(* IEC 61131-3 sources: plc_NativeGateway/src (part 3) *)

(* ---- NG_ReadAck.st ---- *)
FUNCTION_BLOCK NG_ReadAck
VAR_INPUT
    GatewayId : NG_Id;
END_VAR
VAR_IN_OUT
    Doc : NG_Document;
END_VAR
VAR_OUTPUT
    Valid : BOOL;
    MessageId : NG_Id;
    Stored : BOOL;
    Retryable : BOOL;
    Codes : NG_Text;
END_VAR
VAR
    RootFields : NG_AckFields;
    ErrorFields : NG_AckFields;
    t : INT;
    n : INT;
    e : INT;
    count : INT;
    code : NG_Text;
    wire : NG_Text;
END_VAR
Valid := FALSE; MessageId := ''; Stored := FALSE; Retryable := TRUE; Codes := '';
RootFields(Parent:=1,ErrorObject:=FALSE,Doc:=Doc); IF NOT RootFields.Valid THEN RETURN; END_IF;
t := RootFields.Fields[1]; IF (Doc.Tokens[t].Kind<>4) OR (Doc.Tokens[t].Number<>1) THEN RETURN; END_IF;
t := RootFields.Fields[2]; IF (Doc.Tokens[t].Kind<>3) OR (Doc.Tokens[t].Text<>GatewayId) THEN RETURN; END_IF;
t := RootFields.Fields[3];
(* Guard range before conversion. TO_LINT rounds and changes max-safe odd integers. *)
IF Doc.Tokens[t].Kind<>4 THEN RETURN; END_IF;
IF NOT ((Doc.Tokens[t].Number>=0) AND (Doc.Tokens[t].Number<=LREAL#9007199254740991.0)) THEN RETURN; END_IF;
IF Doc.Tokens[t].Number<>TO_LREAL(TRUNC_LINT(Doc.Tokens[t].Number)) THEN RETURN; END_IF;
t := RootFields.Fields[4];
IF (Doc.Tokens[t].Kind<>3) OR (LEN(Doc.Tokens[t].Text)>64) THEN RETURN; END_IF;
MessageId := Doc.Tokens[t].Text; IF NOT NG_ValidId(MessageId) THEN RETURN; END_IF;
t := RootFields.Fields[5]; IF Doc.Tokens[t].Kind<>3 THEN RETURN; END_IF;
IF Doc.Tokens[t].Text='STORED' THEN Stored:=TRUE;
ELSIF Doc.Tokens[t].Text<>'REJECTED' THEN RETURN; END_IF;
n := RootFields.Fields[6]; IF Doc.Tokens[n].Kind<>2 THEN RETURN; END_IF;
e:=n+1; count:=0;
WHILE e<Doc.Tokens[n].NextToken DO
    count:=count+1; IF Stored OR (count>32) THEN RETURN; END_IF;
    ErrorFields(Parent:=e,ErrorObject:=TRUE,Doc:=Doc); IF NOT ErrorFields.Valid THEN RETURN; END_IF;
    t:=ErrorFields.Fields[1]; IF (Doc.Tokens[t].Kind<>3) OR (Doc.Tokens[t].TextLength>256) THEN RETURN; END_IF;
    code:=Doc.Tokens[t].Text; wire:=NG_WireCode(code,FALSE); IF wire<>code THEN RETURN; END_IF;
    IF (code<>'UNKNOWN_CONFIG_VERSION') AND (code<>'RESOURCE_LIMIT') AND (code<>'STORAGE_ERROR') THEN Retryable:=FALSE; END_IF;
    IF LEN(Codes)<200 THEN IF Codes<>'' THEN Codes:=CONCAT(Codes,','); END_IF; Codes:=CONCAT(Codes,code); END_IF;
    t:=ErrorFields.Fields[2]; IF (Doc.Tokens[t].Kind<>3) OR (Doc.Tokens[t].TextLength>512) THEN RETURN; END_IF;
    IF (Doc.Tokens[t].Text<>'') AND (LEFT(Doc.Tokens[t].Text,1)<>'/') THEN RETURN; END_IF;
    t:=ErrorFields.Fields[3]; IF (Doc.Tokens[t].Kind<>3) OR (Doc.Tokens[t].TextLength<1) OR (Doc.Tokens[t].TextLength>256) THEN RETURN; END_IF;
    t:=ErrorFields.Fields[4];
    IF t>0 THEN IF (Doc.Tokens[t].Kind<>3) OR (LEN(Doc.Tokens[t].Text)>64) THEN RETURN; END_IF; wire:=Doc.Tokens[t].Text; IF NOT NG_ValidId(wire) THEN RETURN; END_IF; END_IF;
    t:=ErrorFields.Fields[5];
    IF t>0 THEN IF (Doc.Tokens[t].Kind<>3) OR (LEN(Doc.Tokens[t].Text)>64) THEN RETURN; END_IF; wire:=Doc.Tokens[t].Text; IF NOT NG_ValidId(wire) THEN RETURN; END_IF; END_IF;
    e:=Doc.Tokens[e].NextToken;
END_WHILE;
IF NOT Stored AND (count=0) THEN RETURN; END_IF;
Valid:=TRUE;
END_FUNCTION_BLOCK

(* ---- NG_ReadConfig.st ---- *)
FUNCTION_BLOCK NG_ReadConfig
VAR_INPUT
    Node : INT;
END_VAR
VAR_IN_OUT
    Doc : NG_Document;
    Config : NG_Config;
END_VAR
VAR_OUTPUT
    ErrorText : NG_Text;
END_VAR
VAR
    ReadDevice : NG_ReadDevice;
    Change : NG_EditDevice;
    Device : NG_Device;
    Points : ARRAY[1..32] OF NG_Point;
    t : INT;
    a : INT;
    d : INT;
    r : INT;
    err : NG_Text;
END_VAR
ErrorText := 'SCHEMA_INVALID';
IF NOT NG_Allowed(Node,'|enabled|report|devices|',Doc) THEN RETURN; END_IF;
t := NG_Member(Node,'enabled',Doc);
IF Doc.Tokens[t].Kind <> 5 THEN RETURN; END_IF;
Config.enabled := Doc.Tokens[t].Text = 'true';
r := NG_Member(Node,'report',Doc);
IF NOT NG_Allowed(r,'|batchIntervalMs|maxBatchPoints|',Doc) THEN RETURN; END_IF;
t := NG_Member(r,'batchIntervalMs',Doc);
IF (Doc.Tokens[t].Kind <> 4) OR (Doc.Tokens[t].Number < 1) OR (Doc.Tokens[t].Number > 86400000) OR (Doc.Tokens[t].Number <> TO_LREAL(TO_LINT(Doc.Tokens[t].Number))) THEN RETURN; END_IF;
Config.batchIntervalMs := TO_UDINT(Doc.Tokens[t].Number);
t := NG_Member(r,'maxBatchPoints',Doc);
IF (Doc.Tokens[t].Kind <> 4) OR (Doc.Tokens[t].Number < 1) OR (Doc.Tokens[t].Number > 500) OR (Doc.Tokens[t].Number <> TO_LREAL(TO_LINT(Doc.Tokens[t].Number))) THEN RETURN; END_IF;
Config.maxBatchPoints := TO_UINT(Doc.Tokens[t].Number);
a := NG_Member(Node,'devices',Doc);
IF Doc.Tokens[a].Kind <> 2 THEN RETURN; END_IF;
d := a + 1; Config.DeviceCount := 0; Config.PointCount := 0;
WHILE d < Doc.Tokens[a].NextToken DO
    IF Config.DeviceCount >= 50 THEN ErrorText := 'POINT_LIMIT_EXCEEDED'; RETURN; END_IF;
    ReadDevice(Node := d, Doc := Doc, Device := Device, Points := Points);
    err := ReadDevice.ErrorText;
    IF err <> '' THEN ErrorText := err; RETURN; END_IF;
    Change(DeviceIndex := Config.DeviceCount+1, Remove := FALSE, Replacement := Device, Config := Config, Points := Points);
    IF Change.ErrorText <> '' THEN ErrorText := Change.ErrorText; RETURN; END_IF;
    d := Doc.Tokens[d].NextToken;
END_WHILE;
ErrorText := NG_CheckConfig(Config);
END_FUNCTION_BLOCK

(* ---- NG_ReadDevice.st ---- *)
FUNCTION_BLOCK NG_ReadDevice
VAR_INPUT
    Node : INT;
END_VAR
VAR_IN_OUT
    Doc : NG_Document;
    Device : NG_Device;
    Points : ARRAY[1..32] OF NG_Point;
END_VAR
VAR_OUTPUT
    ErrorText : NG_Text;
END_VAR
VAR
    ReadPoint : NG_ReadPoint;
    t : INT;
    conn : INT;
    pointsNode : INT;
    p : INT;
    err : NG_Text;
END_VAR
ErrorText := '';
IF NOT NG_Allowed(Node,'|deviceId|name|enabled|protocol|connection|points|',Doc) THEN ErrorText := 'SCHEMA_INVALID'; RETURN; END_IF;
t := NG_Member(Node, 'deviceId', Doc);
IF (Doc.Tokens[t].Kind <> 3) OR (LEN(Doc.Tokens[t].Text) < 1) OR (LEN(Doc.Tokens[t].Text) > 64) THEN ErrorText := 'SCHEMA_INVALID'; RETURN; END_IF;
Device.deviceId := Doc.Tokens[t].Text;
t := NG_Member(Node, 'name', Doc);
IF (Doc.Tokens[t].Kind <> 3) OR (LEN(Doc.Tokens[t].Text) < 1) OR (LEN(Doc.Tokens[t].Text) > 128) THEN ErrorText := 'SCHEMA_INVALID'; RETURN; END_IF;
Device.name := Doc.Tokens[t].Text;
t := NG_Member(Node, 'enabled', Doc);
IF (Doc.Tokens[t].Kind <> 5) THEN ErrorText := 'SCHEMA_INVALID'; RETURN; END_IF;
Device.enabled := (Doc.Tokens[t].Text = 'true');
t := NG_Member(Node,'protocol',Doc);
IF (Doc.Tokens[t].Kind <> 3) OR (Doc.Tokens[t].Text <> 'modbus_tcp') THEN ErrorText := 'UNSUPPORTED_PROTOCOL'; RETURN; END_IF;
conn := NG_Member(Node,'connection',Doc);
IF NOT NG_Allowed(conn,'|host|port|unitId|connectTimeoutMs|requestTimeoutMs|retryCount|maxReadRegisters|maxRegisterGap|',Doc) THEN ErrorText := 'SCHEMA_INVALID'; RETURN; END_IF;
t := NG_Member(conn, 'host', Doc);
IF (Doc.Tokens[t].Kind <> 3) OR (LEN(Doc.Tokens[t].Text) < 1) OR (LEN(Doc.Tokens[t].Text) > 253) THEN ErrorText := 'SCHEMA_INVALID'; RETURN; END_IF;
Device.host := Doc.Tokens[t].Text;
t := NG_Member(conn, 'port', Doc);
IF (Doc.Tokens[t].Kind <> 4) OR (Doc.Tokens[t].Number < LREAL#1.0) OR (Doc.Tokens[t].Number > LREAL#65535.0) OR (Doc.Tokens[t].Number <> TO_LREAL(TO_LINT(Doc.Tokens[t].Number))) THEN ErrorText := 'SCHEMA_INVALID'; RETURN; END_IF;
Device.port := TO_UINT(Doc.Tokens[t].Number);
t := NG_Member(conn, 'unitId', Doc);
IF (Doc.Tokens[t].Kind <> 4) OR (Doc.Tokens[t].Number < LREAL#0.0) OR (Doc.Tokens[t].Number > LREAL#255.0) OR (Doc.Tokens[t].Number <> TO_LREAL(TO_LINT(Doc.Tokens[t].Number))) THEN ErrorText := 'SCHEMA_INVALID'; RETURN; END_IF;
Device.unitId := TO_USINT(Doc.Tokens[t].Number);
t := NG_Member(conn, 'connectTimeoutMs', Doc);
IF (Doc.Tokens[t].Kind <> 4) OR (Doc.Tokens[t].Number < LREAL#1.0) OR (Doc.Tokens[t].Number > LREAL#300000.0) OR (Doc.Tokens[t].Number <> TO_LREAL(TO_LINT(Doc.Tokens[t].Number))) THEN ErrorText := 'SCHEMA_INVALID'; RETURN; END_IF;
Device.connectTimeoutMs := TO_UDINT(Doc.Tokens[t].Number);
t := NG_Member(conn, 'requestTimeoutMs', Doc);
IF (Doc.Tokens[t].Kind <> 4) OR (Doc.Tokens[t].Number < LREAL#1.0) OR (Doc.Tokens[t].Number > LREAL#300000.0) OR (Doc.Tokens[t].Number <> TO_LREAL(TO_LINT(Doc.Tokens[t].Number))) THEN ErrorText := 'SCHEMA_INVALID'; RETURN; END_IF;
Device.requestTimeoutMs := TO_UDINT(Doc.Tokens[t].Number);
t := NG_Member(conn, 'retryCount', Doc);
IF (Doc.Tokens[t].Kind <> 4) OR (Doc.Tokens[t].Number < LREAL#0.0) OR (Doc.Tokens[t].Number > LREAL#10.0) OR (Doc.Tokens[t].Number <> TO_LREAL(TO_LINT(Doc.Tokens[t].Number))) THEN ErrorText := 'SCHEMA_INVALID'; RETURN; END_IF;
Device.retryCount := TO_USINT(Doc.Tokens[t].Number);
t := NG_Member(conn, 'maxReadRegisters', Doc);
IF t > 0 THEN
    IF (Doc.Tokens[t].Kind <> 4) OR (Doc.Tokens[t].Number < LREAL#1.0) OR (Doc.Tokens[t].Number > LREAL#125.0) OR (Doc.Tokens[t].Number <> TO_LREAL(TO_LINT(Doc.Tokens[t].Number))) THEN ErrorText := 'SCHEMA_INVALID'; RETURN; END_IF;
    Device.maxReadRegisters := TO_UINT(Doc.Tokens[t].Number);
ELSE
    Device.maxReadRegisters := UINT#0;
END_IF;
t := NG_Member(conn, 'maxRegisterGap', Doc);
IF t > 0 THEN
    IF (Doc.Tokens[t].Kind <> 4) OR (Doc.Tokens[t].Number < LREAL#0.0) OR (Doc.Tokens[t].Number > LREAL#124.0) OR (Doc.Tokens[t].Number <> TO_LREAL(TO_LINT(Doc.Tokens[t].Number))) THEN ErrorText := 'SCHEMA_INVALID'; RETURN; END_IF;
    Device.hasMaxRegisterGap := TRUE;
    Device.maxRegisterGap := TO_UINT(Doc.Tokens[t].Number);
ELSE
    Device.hasMaxRegisterGap := FALSE;
    Device.maxRegisterGap := UINT#0;
END_IF;
pointsNode := NG_Member(Node,'points',Doc);
IF Doc.Tokens[pointsNode].Kind <> 2 THEN ErrorText := 'SCHEMA_INVALID'; RETURN; END_IF;
Device.PointCount := 0; p := pointsNode + 1;
WHILE p < Doc.Tokens[pointsNode].NextToken DO
    IF Device.PointCount >= 32 THEN ErrorText := 'POINT_LIMIT_EXCEEDED'; RETURN; END_IF;
    Device.PointCount := Device.PointCount + 1;
    ReadPoint(Node := p, Doc := Doc, Point := Points[Device.PointCount]);
    err := ReadPoint.ErrorText;
    IF err <> '' THEN ErrorText := err; RETURN; END_IF;
    p := Doc.Tokens[p].NextToken;
END_WHILE;

END_FUNCTION_BLOCK

(* ---- NG_ReadPoint.st ---- *)
FUNCTION_BLOCK NG_ReadPoint
VAR_INPUT
    Node : INT;
END_VAR
VAR_IN_OUT
    Doc : NG_Document;
    Point : NG_Point;
END_VAR
VAR_OUTPUT
    ErrorText : NG_Text;
END_VAR
VAR
    t : INT;
    mb : INT;
END_VAR
ErrorText := '';
IF NOT NG_Allowed(Node,'|pointId|name|enabled|dataType|pollIntervalMs|scale|offset|unit|reportMode|reportIntervalMs|deadband|staleAfterMs|modbus|',Doc) THEN ErrorText := 'SCHEMA_INVALID'; RETURN; END_IF;
t := NG_Member(Node, 'pointId', Doc);
IF (Doc.Tokens[t].Kind <> 3) OR (LEN(Doc.Tokens[t].Text) < 1) OR (LEN(Doc.Tokens[t].Text) > 64) THEN ErrorText := 'SCHEMA_INVALID'; RETURN; END_IF;
Point.pointId := Doc.Tokens[t].Text;
t := NG_Member(Node, 'name', Doc);
IF (Doc.Tokens[t].Kind <> 3) OR (LEN(Doc.Tokens[t].Text) < 1) OR (LEN(Doc.Tokens[t].Text) > 128) THEN ErrorText := 'SCHEMA_INVALID'; RETURN; END_IF;
Point.name := Doc.Tokens[t].Text;
t := NG_Member(Node, 'enabled', Doc);
IF (Doc.Tokens[t].Kind <> 5) THEN ErrorText := 'SCHEMA_INVALID'; RETURN; END_IF;
Point.enabled := (Doc.Tokens[t].Text = 'true');
t := NG_Member(Node, 'dataType', Doc);
IF (Doc.Tokens[t].Kind <> 3) OR (LEN(Doc.Tokens[t].Text) < 1) OR (LEN(Doc.Tokens[t].Text) > 16) THEN ErrorText := 'SCHEMA_INVALID'; RETURN; END_IF;
Point.dataType := Doc.Tokens[t].Text;
t := NG_Member(Node, 'pollIntervalMs', Doc);
IF (Doc.Tokens[t].Kind <> 4) OR (Doc.Tokens[t].Number < LREAL#1.0) OR (Doc.Tokens[t].Number > LREAL#86400000.0) OR (Doc.Tokens[t].Number <> TO_LREAL(TO_LINT(Doc.Tokens[t].Number))) THEN ErrorText := 'SCHEMA_INVALID'; RETURN; END_IF;
Point.pollIntervalMs := TO_UDINT(Doc.Tokens[t].Number);
t := NG_Member(Node, 'scale', Doc);
IF (Doc.Tokens[t].Kind <> 4) OR (Doc.Tokens[t].Number < LREAL#-1.0E+100) OR (Doc.Tokens[t].Number > LREAL#1.0E+100) THEN ErrorText := 'SCHEMA_INVALID'; RETURN; END_IF;
Point.scale := Doc.Tokens[t].Number;
t := NG_Member(Node, 'offset', Doc);
IF (Doc.Tokens[t].Kind <> 4) OR (Doc.Tokens[t].Number < LREAL#-1.0E+100) OR (Doc.Tokens[t].Number > LREAL#1.0E+100) THEN ErrorText := 'SCHEMA_INVALID'; RETURN; END_IF;
Point.offset := Doc.Tokens[t].Number;
t := NG_Member(Node, 'unit', Doc);
IF t > 0 THEN
IF (Doc.Tokens[t].Kind <> 3) OR (LEN(Doc.Tokens[t].Text) < 0) OR (LEN(Doc.Tokens[t].Text) > 32) THEN ErrorText := 'SCHEMA_INVALID'; RETURN; END_IF;
Point.unit := Doc.Tokens[t].Text;
ELSE Point.unit := ''; END_IF;
t := NG_Member(Node, 'reportMode', Doc);
IF (Doc.Tokens[t].Kind <> 3) OR (LEN(Doc.Tokens[t].Text) < 1) OR (LEN(Doc.Tokens[t].Text) > 24) THEN ErrorText := 'SCHEMA_INVALID'; RETURN; END_IF;
Point.reportMode := Doc.Tokens[t].Text;
t := NG_Member(Node, 'reportIntervalMs', Doc);
IF (Doc.Tokens[t].Kind <> 4) OR (Doc.Tokens[t].Number < LREAL#1.0) OR (Doc.Tokens[t].Number > LREAL#86400000.0) OR (Doc.Tokens[t].Number <> TO_LREAL(TO_LINT(Doc.Tokens[t].Number))) THEN ErrorText := 'SCHEMA_INVALID'; RETURN; END_IF;
Point.reportIntervalMs := TO_UDINT(Doc.Tokens[t].Number);
t := NG_Member(Node, 'deadband', Doc);
IF (Doc.Tokens[t].Kind <> 4) OR (Doc.Tokens[t].Number < LREAL#0.0) OR (Doc.Tokens[t].Number > LREAL#1.0E+100) THEN ErrorText := 'SCHEMA_INVALID'; RETURN; END_IF;
Point.deadband := Doc.Tokens[t].Number;
t := NG_Member(Node, 'staleAfterMs', Doc);
IF (Doc.Tokens[t].Kind <> 4) OR (Doc.Tokens[t].Number < LREAL#1.0) OR (Doc.Tokens[t].Number > LREAL#86400000.0) OR (Doc.Tokens[t].Number <> TO_LREAL(TO_LINT(Doc.Tokens[t].Number))) THEN ErrorText := 'SCHEMA_INVALID'; RETURN; END_IF;
Point.staleAfterMs := TO_UDINT(Doc.Tokens[t].Number);
mb := NG_Member(Node,'modbus',Doc);
IF NOT NG_Allowed(mb,'|area|address|byteOrder|',Doc) THEN ErrorText := 'SCHEMA_INVALID'; RETURN; END_IF;
t := NG_Member(mb, 'area', Doc);
IF (Doc.Tokens[t].Kind <> 3) OR (LEN(Doc.Tokens[t].Text) < 1) OR (LEN(Doc.Tokens[t].Text) > 24) THEN ErrorText := 'SCHEMA_INVALID'; RETURN; END_IF;
Point.area := Doc.Tokens[t].Text;
t := NG_Member(mb, 'address', Doc);
IF (Doc.Tokens[t].Kind <> 4) OR (Doc.Tokens[t].Number < LREAL#0.0) OR (Doc.Tokens[t].Number > LREAL#65535.0) OR (Doc.Tokens[t].Number <> TO_LREAL(TO_LINT(Doc.Tokens[t].Number))) THEN ErrorText := 'SCHEMA_INVALID'; RETURN; END_IF;
Point.address := TO_UINT(Doc.Tokens[t].Number);
t := NG_Member(mb, 'byteOrder', Doc);
IF t > 0 THEN
IF (Doc.Tokens[t].Kind <> 3) OR (LEN(Doc.Tokens[t].Text) < 0) OR (LEN(Doc.Tokens[t].Text) > 4) THEN ErrorText := 'SCHEMA_INVALID'; RETURN; END_IF;
Point.byteOrder := Doc.Tokens[t].Text;
ELSE Point.byteOrder := ''; END_IF;
END_FUNCTION_BLOCK

(* ---- NG_ReportPolicy.st ---- *)
FUNCTION_BLOCK NG_ReportPolicy
VAR_INPUT
    DeferCapacity : BOOL;
END_VAR
VAR_IN_OUT
    Buffer : NG_Buffer;
END_VAR
VAR
    Event : NG_CaptureEvent;
    Gap : NG_GapLog;
    AuditDecision : NG_AuditDecision;
    s : UINT;
    p : UINT;
    r : UINT;
    c : UINT;
    n : INT;
    slots : ULINT;
    selected : BOOL;
    present : BOOL;
    reject : BOOL;
    reason : USINT;
END_VAR

(* Atomic RAM admission is this mode's local commit boundary. The copied
   baseline has no dependency on delivery order or subsequent slot reuse. *)
FOR n:=1 TO 64 DO
    IF Buffer.WorkDeadlineUs>0 THEN IF GET_MICROSECONDS(TRUE)+ULINT#70>=Buffer.WorkDeadlineUs THEN EXIT; END_IF; END_IF;
    IF Buffer.IngressCount=0 THEN EXIT; END_IF;
    (* A local whole-batch reclaim may need the next bounded scan. Keep this
       raw event undecided until that reclaim; never wait on SDK/ACK here. *)
    IF DeferCapacity AND (Buffer.FreeHead=0) AND (Buffer.HighSlot>=28800) THEN EXIT; END_IF;
    Event:=Buffer.Ingress[Buffer.Head]; s:=Event.ConfigSlot; p:=Event.PointIndex;
    Buffer.Head:=Buffer.Head MOD 512+1; Buffer.IngressCount:=Buffer.IngressCount-1;
    reject:=FALSE; reason:=0;
    IF (s<>Buffer.ActiveSlot) OR (Event.ConfigGeneration<>Buffer.Configs[s].Generation) OR
       (Event.SamplingGeneration<>Buffer.SamplingGeneration) OR NOT Buffer.Cursors[p].Enabled THEN
        Buffer.UndecidedLostEventsTotal:=NG_SafeAdd(Buffer.UndecidedLostEventsTotal,ULINT#1);
        Buffer.AccountingComplete:=FALSE;
        reason:=2; reject:=TRUE;
    ELSE
        present:=((Event.Flags AND WORD#1)<>WORD#0) AND
                 (((Event.Flags AND WORD#2)<>WORD#0) OR ((Event.Flags AND WORD#8)<>WORD#0));
        IF Buffer.PlatformTime THEN
            present:=present AND Buffer.TimeValid AND (Event.ClockRevision=Buffer.ClockRevision)
                AND ((Event.Flags AND WORD#2)<>WORD#0);
        END_IF;
        IF (Buffer.ReportCursors[p].SamplingGeneration<>Event.SamplingGeneration) OR
           (Buffer.ReportCursors[p].ConfigGeneration<>Event.ConfigGeneration) OR
           (Buffer.ReportCursors[p].ClockRevision<>Event.ClockRevision) OR
           (Buffer.ReportCursors[p].TimePresent<>present) THEN
            slots:=Buffer.Cursors[p].ActivatedMonoMs;
            IF (Buffer.ReportCursors[p].ConfigGeneration=Event.ConfigGeneration) AND
               ((Buffer.ReportCursors[p].TimePresent<>present) OR (Buffer.ReportCursors[p].ClockRevision<>Event.ClockRevision)) THEN
                slots:=Buffer.Cursors[p].NextDueMonoMs;
                IF Event.Kind=1 THEN slots:=Event.NominalDueMonoMs; END_IF;
            END_IF;
            Buffer.ReportCursors[p].SamplingGeneration:=Event.SamplingGeneration;
            Buffer.ReportCursors[p].ConfigGeneration:=Event.ConfigGeneration;
            Buffer.ReportCursors[p].ClockRevision:=Event.ClockRevision;
            Buffer.ReportCursors[p].TimePresent:=present;
            Buffer.ReportCursors[p].HasBaseline:=FALSE;
            Buffer.ReportCursors[p].NextDue:=slots;
        END_IF;
        selected:=NOT Buffer.ReportCursors[p].HasBaseline OR (Buffer.ReportCursors[p].Quality<>Event.Quality);
        IF Buffer.ReportCursors[p].HasBaseline AND (Event.Quality=2) AND (Buffer.ReportCursors[p].Quality=2) AND
           (Buffer.Configs[s].Config.Points[p].reportMode<>'cyclic') THEN
            IF Buffer.Configs[s].Config.Points[p].dataType='bool' THEN
                selected:=selected OR ((Event.Value=LREAL#0.0)<>(Buffer.ReportCursors[p].Value=LREAL#0.0));
            ELSE selected:=selected OR (ABS(Event.Value-Buffer.ReportCursors[p].Value)>Buffer.Configs[s].Config.Points[p].deadband); END_IF;
        END_IF;
        IF (Event.Kind=1) AND (Buffer.Configs[s].Config.Points[p].reportMode<>'change') AND
           (Event.NominalDueMonoMs>=Buffer.ReportCursors[p].NextDue) THEN
            slots:=(Event.NominalDueMonoMs-Buffer.ReportCursors[p].NextDue)/TO_ULINT(Buffer.Configs[s].Config.Points[p].reportIntervalMs)+1;
            Buffer.MissedReportSlotsTotal:=NG_SafeAdd(Buffer.MissedReportSlotsTotal,slots-1);
            Buffer.ReportCursors[p].NextDue:=Buffer.ReportCursors[p].NextDue+slots*TO_ULINT(Buffer.Configs[s].Config.Points[p].reportIntervalMs);
            selected:=TRUE;
        END_IF;
        IF NOT selected THEN
            Buffer.PolicyFilteredEventsTotal:=NG_SafeAdd(Buffer.PolicyFilteredEventsTotal,ULINT#1); reject:=TRUE;
        ELSE
            Buffer.EligibleEventsTotal:=NG_SafeAdd(Buffer.EligibleEventsTotal,ULINT#1);
            IF NOT present THEN
                Buffer.TimeInvalidEventsTotal:=NG_SafeAdd(Buffer.TimeInvalidEventsTotal,ULINT#1); reason:=4; reject:=TRUE;
            ELSIF (Buffer.FreeHead=0) AND (Buffer.HighSlot>=28800) THEN
                Buffer.EnqueueRejectedAttemptsTotal:=NG_SafeAdd(Buffer.EnqueueRejectedAttemptsTotal,ULINT#1); reason:=5; reject:=TRUE;
            END_IF;
            IF reject THEN Buffer.KnownUnsentEventsTotal:=NG_SafeAdd(Buffer.KnownUnsentEventsTotal,ULINT#1); END_IF;
        END_IF;
    END_IF;
    IF reject THEN
        c:=1;
        IF reason=2 THEN c:=4; ELSIF reason<>0 THEN c:=3; END_IF;
        AuditDecision(SampleSeq:=Event.SampleSeq,Decision:=TO_USINT(c),Reason:=reason,Buffer:=Buffer);
        IF reason<>0 THEN Gap(Reason:=reason,Event:=Event,Buffer:=Buffer); END_IF;
        Buffer.Configs[s].References:=Buffer.Configs[s].References-1;
    ELSE
        IF Buffer.FreeHead<>0 THEN r:=Buffer.FreeHead; Buffer.FreeHead:=Buffer.FreeSlots[r];
        ELSE Buffer.HighSlot:=Buffer.HighSlot+1; r:=Buffer.HighSlot; END_IF;
        IF Buffer.RecordGenerations[r]=UDINT#4294967295 THEN Buffer.CaptureStopped:=TRUE;
            Buffer.KnownUnsentEventsTotal:=NG_SafeAdd(Buffer.KnownUnsentEventsTotal,ULINT#1);
            Gap(Reason:=USINT#5,Event:=Event,Buffer:=Buffer); Buffer.Configs[s].References:=Buffer.Configs[s].References-1;
            AuditDecision(SampleSeq:=Event.SampleSeq,Decision:=USINT#3,Reason:=USINT#5,Buffer:=Buffer);
        ELSE
            Buffer.RecordGenerations[r]:=Buffer.RecordGenerations[r]+1;
            Buffer.Records[r]:=Event; Buffer.RecordStates[r]:=1; Buffer.FreeSlots[r]:=0;
            Buffer.LastAdmittedSeq:=MAX(Buffer.LastAdmittedSeq,Event.SampleSeq);
            AuditDecision(SampleSeq:=Event.SampleSeq,Decision:=USINT#2,Reason:=USINT#0,Buffer:=Buffer);
            Buffer.OwnedCount:=Buffer.OwnedCount+1;
            c:=2; IF Event.SampleSeq<=Buffer.Watermark THEN c:=1; END_IF;
            IF Buffer.QueueHead[c]=0 THEN Buffer.QueueHead[c]:=r; ELSE Buffer.FreeSlots[Buffer.QueueTail[c]]:=r; END_IF;
            Buffer.QueueTail[c]:=r;
            IF Event.SampleSeq>Buffer.ReportCursors[p].LastSeq THEN
                Buffer.ReportCursors[p].LastSeq:=Event.SampleSeq; Buffer.ReportCursors[p].Value:=Event.Value;
                Buffer.ReportCursors[p].Quality:=Event.Quality; Buffer.ReportCursors[p].HasBaseline:=TRUE;
            END_IF;
        END_IF;
    END_IF;
END_FOR;
END_FUNCTION_BLOCK

(* ---- NG_Resources.st ---- *)
FUNCTION_BLOCK NG_Resources
VAR_INPUT
    NowMs : ULINT;
END_VAR
VAR_OUTPUT
    Changed : BOOL;
    MemoryValid : BOOL;
    CpuValid : BOOL;
    ProcessValid : BOOL;
    TotalKiB : ULINT;
    AvailableKiB : ULINT;
    RssKiB : ULINT;
    CpuPermille : UDINT;
    ProcessName : STRING[64];
    ErrorText : NG_Text;
END_VAR
VAR
    OpenFile : FILE_OPEN;
    ReadFile : FILE_READ;
    CloseFile : FILE_CLOSE;
    Convert : BUF_TO_STRING;
    Name : STRING;
    Bytes : NG_ProcBytes;
    Text : NG_ProcText;
    Stage : INT;
    FileIndex : INT := 1;
    Handle : UINT;
    Count : UDINT;
    NextRead : ULINT;
    p : INT;
    c : INT;
    n : INT;
    start : INT;
    token : ULINT;
    total : ULINT;
    idle : ULINT;
    PrevTotal : ULINT;
    PrevIdle : ULINT;
    HasDigit : BOOL;
    ProcFailed : BOOL;
END_VAR
Changed := FALSE;
CASE FileIndex OF
1: Name := '/proc/meminfo';
2: Name := '/proc/stat';
3: Name := '/proc/self/status';
END_CASE;
OpenFile(Execute := Stage=10, Name := Name);
ReadFile(Execute := Stage=20, Handle := Handle, MaxLength := UDINT#8191, Buffer := Bytes);
CloseFile(Execute := Stage=30, Handle := Handle);
Convert(REQ := Stage=40, BUF_FORMAT := FALSE, BUF_OFFS := 0, BUF_CNT := TO_INT(Count), BUFFER := Bytes, DST := Text);
CASE Stage OF
0:
    IF NowMs >= NextRead THEN FileIndex := 1; ErrorText := ''; ProcFailed := FALSE; Stage := 10; END_IF;
10:
    IF OpenFile.Error THEN ProcFailed := TRUE; Stage := 80;
    ELSIF OpenFile.Done THEN Handle := OpenFile.Handle; Stage := 20; END_IF;
20:
    IF ReadFile.Error OR ReadFile.Done THEN Count := ReadFile.LengthRead; ProcFailed := Count=0; Stage := 30; END_IF;
30:
    IF CloseFile.Done OR CloseFile.Error THEN IF CloseFile.Error OR ProcFailed THEN Stage := 80; ELSE Stage := 40; END_IF; END_IF;
40:
    IF Convert.ERROR THEN ProcFailed := TRUE; Stage := 80;
    ELSIF Convert.DONE THEN
        CASE FileIndex OF
        1:
            TotalKiB := NG_ProcNumber(Text,'MemTotal:'); AvailableKiB := NG_ProcNumber(Text,'MemAvailable:');
            IF AvailableKiB=0 THEN AvailableKiB := NG_ProcNumber(Text,'MemFree:')+NG_ProcNumber(Text,'Buffers:')+NG_ProcNumber(Text,'Cached:'); END_IF;
            MemoryValid := TotalKiB > 0;
        2:
            total := 0; idle := 0; n := 0; token := 0; HasDigit := FALSE;
            p := FIND(Text,'cpu ');
            IF p > 0 THEN
                p := p+4;
                WHILE p <= LEN(Text) DO
                    c := GET_CHAR(Text,p);
                    IF (c>=48) AND (c<=57) THEN token := token*10+TO_ULINT(c-48); HasDigit := TRUE;
                    ELSE
                        IF HasDigit THEN
                            n := n+1; IF n <= 8 THEN total := total+token; END_IF;
                            IF (n=4) OR (n=5) THEN idle := idle+token; END_IF;
                            token := 0; HasDigit := FALSE;
                        END_IF;
                        IF (c=10) OR (n>=8) THEN EXIT; END_IF;
                    END_IF;
                    p := p+1;
                END_WHILE;
                IF (PrevTotal > 0) AND (total > PrevTotal) AND (idle >= PrevIdle) THEN
                    CpuPermille := TO_UDINT((total-PrevTotal-(idle-PrevIdle))*1000/(total-PrevTotal)); CpuValid := TRUE;
                END_IF;
                PrevTotal := total; PrevIdle := idle;
            END_IF;
        3:
            RssKiB := NG_ProcNumber(Text,'VmRSS:'); ProcessValid := RssKiB > 0;
            start := FIND(Text,'Name:');
            IF start > 0 THEN
                start := start+5;
                WHILE start <= LEN(Text) DO c := GET_CHAR(Text,start); IF (c<>32) AND (c<>9) THEN EXIT; END_IF; start := start+1; END_WHILE;
                p := start;
                WHILE p <= LEN(Text) DO IF GET_CHAR(Text,p)=10 THEN EXIT; END_IF; p := p+1; END_WHILE;
                IF p > start THEN ProcessName := MID(Text,MIN(63,p-start),start); END_IF;
            END_IF;
        END_CASE;
        Stage := 80;
    END_IF;
80:
    IF ProcFailed THEN
        ErrorText := CONCAT('PROC_READ_FAILED:',TO_STRING(FileIndex,'{0:d}'));
        CASE FileIndex OF 1: MemoryValid := FALSE; 2: CpuValid := FALSE; 3: ProcessValid := FALSE; END_CASE;
    END_IF;
    ProcFailed := FALSE;
    IF FileIndex < 3 THEN FileIndex := FileIndex+1; Stage := 10;
    ELSE Changed := TRUE; NextRead := NowMs+10000; Stage := 0; END_IF;
END_CASE;
END_FUNCTION_BLOCK

(* ---- NG_SameConfig.st ---- *)
FUNCTION_BLOCK NG_SameConfig
VAR_OUTPUT
    Equal : BOOL;
END_VAR
VAR_IN_OUT
    A : NG_Config;
    B : NG_Config;
END_VAR
VAR
    i : INT;
END_VAR
Equal := FALSE;
IF (A.Version<>B.Version) OR (A.MessageId<>B.MessageId) OR (A.enabled<>B.enabled) OR
   (A.batchIntervalMs<>B.batchIntervalMs) OR (A.maxBatchPoints<>B.maxBatchPoints) OR
   (A.DeviceCount<>B.DeviceCount) OR (A.PointCount<>B.PointCount) THEN RETURN; END_IF;
FOR i:=1 TO A.DeviceCount DO
    IF (A.Devices[i].deviceId<>B.Devices[i].deviceId) OR (A.Devices[i].name<>B.Devices[i].name) OR
       (A.Devices[i].enabled<>B.Devices[i].enabled) OR (A.Devices[i].host<>B.Devices[i].host) OR
       (A.Devices[i].port<>B.Devices[i].port) OR (A.Devices[i].unitId<>B.Devices[i].unitId) OR
       (A.Devices[i].connectTimeoutMs<>B.Devices[i].connectTimeoutMs) OR
       (A.Devices[i].requestTimeoutMs<>B.Devices[i].requestTimeoutMs) OR
       (A.Devices[i].retryCount<>B.Devices[i].retryCount) OR
       (A.Devices[i].maxReadRegisters<>B.Devices[i].maxReadRegisters) OR
       (A.Devices[i].hasMaxRegisterGap<>B.Devices[i].hasMaxRegisterGap) OR
       (A.Devices[i].maxRegisterGap<>B.Devices[i].maxRegisterGap) OR
       (A.Devices[i].PointStart<>B.Devices[i].PointStart) OR (A.Devices[i].PointCount<>B.Devices[i].PointCount) THEN RETURN; END_IF;
END_FOR;
FOR i:=1 TO A.PointCount DO
    IF (A.Points[i].pointId<>B.Points[i].pointId) OR (A.Points[i].name<>B.Points[i].name) OR
       (A.Points[i].enabled<>B.Points[i].enabled) OR (A.Points[i].dataType<>B.Points[i].dataType) OR
       (A.Points[i].pollIntervalMs<>B.Points[i].pollIntervalMs) OR (A.Points[i].scale<>B.Points[i].scale) OR
       (A.Points[i].offset<>B.Points[i].offset) OR (A.Points[i].unit<>B.Points[i].unit) OR
       (A.Points[i].reportMode<>B.Points[i].reportMode) OR (A.Points[i].reportIntervalMs<>B.Points[i].reportIntervalMs) OR
       (A.Points[i].deadband<>B.Points[i].deadband) OR (A.Points[i].staleAfterMs<>B.Points[i].staleAfterMs) OR
       (A.Points[i].area<>B.Points[i].area) OR (A.Points[i].address<>B.Points[i].address) OR
       (A.Points[i].byteOrder<>B.Points[i].byteOrder) THEN RETURN; END_IF;
END_FOR;
Equal := TRUE;
END_FUNCTION_BLOCK

(* ---- NG_SHA256.st ---- *)
FUNCTION_BLOCK NG_SHA256
VAR_INPUT
    Execute : BOOL;
    Length : UDINT;
END_VAR
VAR_IN_OUT
    Buffer : NG_Bytes;
END_VAR
VAR_OUTPUT
    Busy : BOOL;
    Done : BOOL;
    Digest : STRING[64];
END_VAR
VAR
    Prev : BOOL;
    Block : UDINT;
    Blocks : UDINT;
    Offset : UDINT;
    i : INT;
    j : INT;
    n : INT;
    v : DWORD;
    a : DWORD;
    b : DWORD;
    c : DWORD;
    d : DWORD;
    e : DWORD;
    f : DWORD;
    g : DWORD;
    h : DWORD;
    s0 : DWORD;
    s1 : DWORD;
    t1 : DWORD;
    t2 : DWORD;
    Hs : ARRAY[0..7] OF DWORD;
    W : ARRAY[0..63] OF DWORD;
    K : ARRAY[0..63] OF DWORD := [16#428A2F98,16#71374491,16#B5C0FBCF,16#E9B5DBA5,16#3956C25B,16#59F111F1,16#923F82A4,16#AB1C5ED5,16#D807AA98,16#12835B01,16#243185BE,16#550C7DC3,16#72BE5D74,16#80DEB1FE,16#9BDC06A7,16#C19BF174,16#E49B69C1,16#EFBE4786,16#0FC19DC6,16#240CA1CC,16#2DE92C6F,16#4A7484AA,16#5CB0A9DC,16#76F988DA,16#983E5152,16#A831C66D,16#B00327C8,16#BF597FC7,16#C6E00BF3,16#D5A79147,16#06CA6351,16#14292967,16#27B70A85,16#2E1B2138,16#4D2C6DFC,16#53380D13,16#650A7354,16#766A0ABB,16#81C2C92E,16#92722C85,16#A2BFE8A1,16#A81A664B,16#C24B8B70,16#C76C51A3,16#D192E819,16#D6990624,16#F40E3585,16#106AA070,16#19A4C116,16#1E376C08,16#2748774C,16#34B0BCB5,16#391C0CB3,16#4ED8AA4A,16#5B9CCA4F,16#682E6FF3,16#748F82EE,16#78A5636F,16#84C87814,16#8CC70208,16#90BEFFFA,16#A4506CEB,16#BEF9A3F7,16#C67178F2];
END_VAR
IF Execute AND NOT Prev AND NOT Busy THEN
    Hs[0] := 16#6A09E667; Hs[1] := 16#BB67AE85; Hs[2] := 16#3C6EF372; Hs[3] := 16#A54FF53A;
    Hs[4] := 16#510E527F; Hs[5] := 16#9B05688C; Hs[6] := 16#1F83D9AB; Hs[7] := 16#5BE0CD19;
    Block := 0; Blocks := (Length + 72) / 64; Busy := TRUE; Done := FALSE; Digest := '';
END_IF;
Prev := Execute;
IF NOT Busy THEN RETURN; END_IF;
FOR n := 1 TO 8 DO
    FOR i := 0 TO 15 DO
        W[i] := 0;
        FOR j := 0 TO 3 DO
            Offset := Block*64 + TO_UDINT(i*4+j);
            IF Offset < Length THEN v := TO_DWORD(Buffer[Offset]);
            ELSIF Offset = Length THEN v := DWORD#16#80;
            ELSIF Offset >= Blocks*64-8 THEN v := TO_DWORD(SHR(TO_LWORD(TO_ULINT(Length)*ULINT#8),TO_UINT((Blocks*64-1-Offset)*8)) AND LWORD#255);
            ELSE v := 0; END_IF;
            W[i] := SHL(W[i],8) OR v;
        END_FOR;
    END_FOR;
    FOR i := 16 TO 63 DO
        s0 := ROR(W[i-15],7) XOR ROR(W[i-15],18) XOR SHR(W[i-15],3);
        s1 := ROR(W[i-2],17) XOR ROR(W[i-2],19) XOR SHR(W[i-2],10);
        W[i] := NG_Add4(W[i-16],s0,W[i-7],s1);
    END_FOR;
    a := Hs[0]; b := Hs[1]; c := Hs[2]; d := Hs[3]; e := Hs[4]; f := Hs[5]; g := Hs[6]; h := Hs[7];
    FOR i := 0 TO 63 DO
        s1 := ROR(e,6) XOR ROR(e,11) XOR ROR(e,25);
        t1 := NG_Add4(h,s1,(e AND f) XOR ((NOT e) AND g),K[i]);
        t1 := NG_Add4(t1,W[i],DWORD#0,DWORD#0);
        s0 := ROR(a,2) XOR ROR(a,13) XOR ROR(a,22);
        t2 := NG_Add4(s0,(a AND b) XOR (a AND c) XOR (b AND c),DWORD#0,DWORD#0);
        h := g; g := f; f := e; e := NG_Add4(d,t1,DWORD#0,DWORD#0);
        d := c; c := b; b := a; a := NG_Add4(t1,t2,DWORD#0,DWORD#0);
    END_FOR;
    Hs[0] := NG_Add4(Hs[0],a,DWORD#0,DWORD#0); Hs[1] := NG_Add4(Hs[1],b,DWORD#0,DWORD#0);
    Hs[2] := NG_Add4(Hs[2],c,DWORD#0,DWORD#0); Hs[3] := NG_Add4(Hs[3],d,DWORD#0,DWORD#0);
    Hs[4] := NG_Add4(Hs[4],e,DWORD#0,DWORD#0); Hs[5] := NG_Add4(Hs[5],f,DWORD#0,DWORD#0);
    Hs[6] := NG_Add4(Hs[6],g,DWORD#0,DWORD#0); Hs[7] := NG_Add4(Hs[7],h,DWORD#0,DWORD#0);
    Block := Block + 1;
    IF Block >= Blocks THEN
        FOR i := 0 TO 7 DO Digest := CONCAT(Digest,TO_STRING(Hs[i],'{0:x8}')); END_FOR;
        Busy := FALSE; Done := TRUE; EXIT;
    END_IF;
END_FOR;
END_FUNCTION_BLOCK

(* ---- NG_SourceResult.st ---- *)
FUNCTION_BLOCK NG_SourceResult
VAR_INPUT
    Index : UINT;
    Value : LREAL;
    Quality : STRING[24];
    NowMs : ULINT;
    UnixMs : ULINT;
    NominalDueMs : ULINT;
    ConfigSlot : UINT;
    ConfigGeneration : UDINT;
    SamplingGeneration : ULINT;
END_VAR
VAR_OUTPUT
    Accepted : BOOL;
END_VAR
VAR_IN_OUT
    Samples : ARRAY[1..320] OF NG_Sample;
    Buffer : NG_Buffer;
END_VAR
VAR
    Core : NG_SourceResultCore;
END_VAR
(* Bind each bounded source/sample/deadline once for the final physical result. *)
Accepted:=FALSE;
IF (Index<1) OR (Index>320) THEN RETURN; END_IF;
Core(Index:=Index,Value:=Value,Quality:=Quality,NowMs:=NowMs,UnixMs:=UnixMs,NominalDueMs:=NominalDueMs,ConfigSlot:=ConfigSlot,ConfigGeneration:=ConfigGeneration,SamplingGeneration:=SamplingGeneration,Cursor:=Buffer.Cursors[Index],Sample:=Samples[Index],StaleDue:=Buffer.SourceStaleDue[Index],Buffer:=Buffer);
Accepted:=Core.Accepted;
END_FUNCTION_BLOCK

(* ---- NG_SourceResultCore.st ---- *)
FUNCTION_BLOCK NG_SourceResultCore
VAR_INPUT
    Index : UINT;
    Value : LREAL;
    Quality : STRING[24];
    NowMs : ULINT;
    UnixMs : ULINT;
    NominalDueMs : ULINT;
    ConfigSlot : UINT;
    ConfigGeneration : UDINT;
    SamplingGeneration : ULINT;
END_VAR
VAR_OUTPUT
    Accepted : BOOL;
END_VAR
VAR_IN_OUT
    Cursor : NG_SourceCursor;
    Sample : NG_Sample;
    StaleDue : ULINT;
    Buffer : NG_Buffer;
END_VAR
VAR
    Capture : NG_Capture;
    code : USINT;
    text : STRING[24];
END_VAR
Accepted:=FALSE;
IF (Index<1) OR (Index>320) OR (ConfigSlot=0) OR (ConfigSlot>4) THEN RETURN; END_IF;
IF (ConfigSlot<>Buffer.ActiveSlot) OR (Buffer.Configs[ConfigSlot].Generation<>ConfigGeneration) OR
   (Buffer.SamplingGeneration<>SamplingGeneration) OR NOT Cursor.Enabled THEN
    Buffer.CancelledReadsTotal:=NG_SafeAdd(Buffer.CancelledReadsTotal,ULINT#1);
    Buffer.CancellationReason:=2; RETURN;
END_IF;
IF NowMs<NominalDueMs THEN Buffer.CaptureStopped:=TRUE; RETURN; END_IF;
text:=Quality;
IF (text='GOOD') AND NOT (ABS(Value)<=LREAL#1.7976931348623157E308) THEN text:='BAD_DECODE'; END_IF;
code:=NG_QualityCode(text);
Capture(PointIndex:=Index, Kind:=USINT#1, Quality:=code, Value:=Value, NowMs:=NowMs, NominalDueMs:=NominalDueMs, SystemUtcMs:=UnixMs, Buffer:=Buffer);
    Accepted:=Capture.Accepted;
Cursor.LastPhysicalMonoMs:=NowMs; Cursor.HasPhysical:=TRUE;
Cursor.Quality:=code;
(* A final result extends this source's liveness. Keeping an earlier global
   deadline is safe; the due sweep recomputes the minimum before emitting stale. *)
StaleDue:=0;
IF code<>3 THEN
    StaleDue:=NowMs+TO_ULINT(Buffer.Configs[ConfigSlot].Config.Points[Index].staleAfterMs);
    IF StaleDue<Buffer.StaleCheckAt THEN Buffer.StaleCheckAt:=StaleDue; END_IF;
END_IF;
Sample.Quality:=text; Sample.Timestamp:=UnixMs; Sample.Fresh:=TRUE;
IF text='GOOD' THEN Sample.Value:=Value; Sample.LastGoodMs:=NowMs; END_IF;
Sample.NextPollMs:=Cursor.NextDueMonoMs;
END_FUNCTION_BLOCK

(* ---- NG_SourceState.st ---- *)
FUNCTION_BLOCK NG_SourceState
VAR_INPUT
    Index : UINT;
    Enabled : BOOL;
    NowMs : ULINT;
    UnixMs : ULINT;
    StaleAfterMs : UDINT;
    CheckStale : BOOL;
END_VAR
VAR_OUTPUT
    Accepted : BOOL;
END_VAR
VAR_IN_OUT
    Samples : ARRAY[1..320] OF NG_Sample;
    Buffer : NG_Buffer;
END_VAR
VAR
    Core : NG_SourceStateCore;
END_VAR
(* Bind each bounded source/sample reference once. Repeated field updates in
   Core avoid dozens of generated array-bound helper calls per activation. *)
Accepted:=FALSE;
IF (Index<1) OR (Index>320) THEN RETURN; END_IF;
Core(Index:=Index,Enabled:=Enabled,NowMs:=NowMs,UnixMs:=UnixMs,
    StaleAfterMs:=StaleAfterMs,CheckStale:=CheckStale,
    Cursor:=Buffer.Cursors[Index],Sample:=Samples[Index],Buffer:=Buffer);
Accepted:=Core.Accepted;
END_FUNCTION_BLOCK

(* ---- NG_SourceStateCore.st ---- *)
FUNCTION_BLOCK NG_SourceStateCore
VAR_INPUT
    Index : UINT;
    Enabled : BOOL;
    NowMs : ULINT;
    UnixMs : ULINT;
    StaleAfterMs : UDINT;
    CheckStale : BOOL;
END_VAR
VAR_OUTPUT
    Accepted : BOOL;
END_VAR
VAR_IN_OUT
    Cursor : NG_SourceCursor;
    Sample : NG_Sample;
    Buffer : NG_Buffer;
END_VAR
VAR
    Capture : NG_CaptureCore;
    start : ULINT;
END_VAR

Accepted:=FALSE;
IF (Index<1) OR (Index>320) THEN RETURN; END_IF;
IF NOT Enabled THEN Cursor.Enabled:=FALSE; Buffer.SourceStaleDue[Index]:=0; RETURN; END_IF;
IF (Cursor.Generation<>Buffer.SamplingGeneration) OR NOT Cursor.Enabled THEN
    Cursor.Generation:=Buffer.SamplingGeneration; Cursor.Enabled:=TRUE;
    Cursor.ActivatedMonoMs:=NowMs; Cursor.LastPhysicalMonoMs:=0;
    Cursor.HasPhysical:=FALSE; Cursor.HasPhysicalUtc:=FALSE;
    Cursor.NextDueMonoMs:=NowMs; Cursor.Quality:=1;
    Buffer.SourceStaleDue[Index]:=NowMs+TO_ULINT(StaleAfterMs);
    IF Buffer.SourceStaleDue[Index]<Buffer.StaleCheckAt THEN Buffer.StaleCheckAt:=Buffer.SourceStaleDue[Index]; END_IF;
    Sample.Quality:='UNKNOWN'; Sample.Timestamp:=UnixMs; Sample.Fresh:=TRUE;
    Sample.NextPollMs:=NowMs;
    Capture(PointIndex:=Index, Kind:=USINT#2, Quality:=USINT#1, Value:=LREAL#0.0, NowMs:=NowMs, NominalDueMs:=ULINT#0, SystemUtcMs:=UnixMs, Cursor:=Cursor, Buffer:=Buffer);
    Accepted:=Capture.Accepted;
END_IF;
IF NOT CheckStale THEN RETURN; END_IF;
start:=Cursor.ActivatedMonoMs;
IF Cursor.HasPhysical THEN start:=Cursor.LastPhysicalMonoMs; END_IF;
IF (NowMs>=start) AND (NowMs-start>=TO_ULINT(StaleAfterMs)) AND (Cursor.Quality<>3) THEN
    Cursor.Quality:=3; Sample.Quality:='STALE';
    Buffer.SourceStaleDue[Index]:=0;
    Sample.Timestamp:=UnixMs; Sample.Fresh:=TRUE;
    Capture(PointIndex:=Index, Kind:=USINT#2, Quality:=USINT#3, Value:=LREAL#0.0, NowMs:=NowMs, NominalDueMs:=ULINT#0, SystemUtcMs:=UnixMs, Cursor:=Cursor, Buffer:=Buffer);
    Accepted:=Capture.Accepted;
END_IF;
END_FUNCTION_BLOCK

(* ---- NG_StorageHash.st ---- *)
FUNCTION_BLOCK NG_StorageHash
VAR_INPUT
    Execute : BOOL;
    Length : UDINT;
END_VAR
VAR_IN_OUT
    Buffer : NG_StorageBytes;
END_VAR
VAR_OUTPUT
    Busy : BOOL;
    Done : BOOL;
    Digest : STRING[64];
END_VAR
VAR
    Prev : BOOL;
    Block : UDINT;
    Blocks : UDINT;
    Offset : UDINT;
    i : INT;
    j : INT;
    n : INT;
    v : DWORD;
    a : DWORD;
    b : DWORD;
    c : DWORD;
    d : DWORD;
    e : DWORD;
    f : DWORD;
    g : DWORD;
    h : DWORD;
    s0 : DWORD;
    s1 : DWORD;
    t1 : DWORD;
    t2 : DWORD;
    Hs : ARRAY[0..7] OF DWORD;
    W : ARRAY[0..63] OF DWORD;
    K : ARRAY[0..63] OF DWORD := [16#428A2F98,16#71374491,16#B5C0FBCF,16#E9B5DBA5,16#3956C25B,16#59F111F1,16#923F82A4,16#AB1C5ED5,16#D807AA98,16#12835B01,16#243185BE,16#550C7DC3,16#72BE5D74,16#80DEB1FE,16#9BDC06A7,16#C19BF174,16#E49B69C1,16#EFBE4786,16#0FC19DC6,16#240CA1CC,16#2DE92C6F,16#4A7484AA,16#5CB0A9DC,16#76F988DA,16#983E5152,16#A831C66D,16#B00327C8,16#BF597FC7,16#C6E00BF3,16#D5A79147,16#06CA6351,16#14292967,16#27B70A85,16#2E1B2138,16#4D2C6DFC,16#53380D13,16#650A7354,16#766A0ABB,16#81C2C92E,16#92722C85,16#A2BFE8A1,16#A81A664B,16#C24B8B70,16#C76C51A3,16#D192E819,16#D6990624,16#F40E3585,16#106AA070,16#19A4C116,16#1E376C08,16#2748774C,16#34B0BCB5,16#391C0CB3,16#4ED8AA4A,16#5B9CCA4F,16#682E6FF3,16#748F82EE,16#78A5636F,16#84C87814,16#8CC70208,16#90BEFFFA,16#A4506CEB,16#BEF9A3F7,16#C67178F2];
END_VAR
IF Execute AND NOT Prev AND NOT Busy THEN
    Hs[0] := 16#6A09E667; Hs[1] := 16#BB67AE85; Hs[2] := 16#3C6EF372; Hs[3] := 16#A54FF53A;
    Hs[4] := 16#510E527F; Hs[5] := 16#9B05688C; Hs[6] := 16#1F83D9AB; Hs[7] := 16#5BE0CD19;
    Block := 0; Blocks := (Length + 72) / 64; Busy := TRUE; Done := FALSE; Digest := '';
END_IF;
Prev := Execute;
IF NOT Busy THEN RETURN; END_IF;
FOR n := 1 TO 16 DO
    FOR i := 0 TO 15 DO
        W[i] := 0;
        FOR j := 0 TO 3 DO
            Offset := Block*64 + TO_UDINT(i*4+j);
            IF Offset < Length THEN v := TO_DWORD(Buffer[Offset]);
            ELSIF Offset = Length THEN v := DWORD#16#80;
            ELSIF Offset >= Blocks*64-8 THEN v := TO_DWORD(SHR(TO_LWORD(TO_ULINT(Length)*ULINT#8),TO_UINT((Blocks*64-1-Offset)*8)) AND LWORD#255);
            ELSE v := 0; END_IF;
            W[i] := SHL(W[i],8) OR v;
        END_FOR;
    END_FOR;
    FOR i := 16 TO 63 DO
        s0 := ROR(W[i-15],7) XOR ROR(W[i-15],18) XOR SHR(W[i-15],3);
        s1 := ROR(W[i-2],17) XOR ROR(W[i-2],19) XOR SHR(W[i-2],10);
        W[i] := NG_Add4(W[i-16],s0,W[i-7],s1);
    END_FOR;
    a := Hs[0]; b := Hs[1]; c := Hs[2]; d := Hs[3]; e := Hs[4]; f := Hs[5]; g := Hs[6]; h := Hs[7];
    FOR i := 0 TO 63 DO
        s1 := ROR(e,6) XOR ROR(e,11) XOR ROR(e,25);
        t1 := NG_Add4(h,s1,(e AND f) XOR ((NOT e) AND g),K[i]);
        t1 := NG_Add4(t1,W[i],DWORD#0,DWORD#0);
        s0 := ROR(a,2) XOR ROR(a,13) XOR ROR(a,22);
        t2 := NG_Add4(s0,(a AND b) XOR (a AND c) XOR (b AND c),DWORD#0,DWORD#0);
        h := g; g := f; f := e; e := NG_Add4(d,t1,DWORD#0,DWORD#0);
        d := c; c := b; b := a; a := NG_Add4(t1,t2,DWORD#0,DWORD#0);
    END_FOR;
    Hs[0] := NG_Add4(Hs[0],a,DWORD#0,DWORD#0); Hs[1] := NG_Add4(Hs[1],b,DWORD#0,DWORD#0);
    Hs[2] := NG_Add4(Hs[2],c,DWORD#0,DWORD#0); Hs[3] := NG_Add4(Hs[3],d,DWORD#0,DWORD#0);
    Hs[4] := NG_Add4(Hs[4],e,DWORD#0,DWORD#0); Hs[5] := NG_Add4(Hs[5],f,DWORD#0,DWORD#0);
    Hs[6] := NG_Add4(Hs[6],g,DWORD#0,DWORD#0); Hs[7] := NG_Add4(Hs[7],h,DWORD#0,DWORD#0);
    Block := Block + 1;
    IF Block >= Blocks THEN
        FOR i := 0 TO 7 DO Digest := CONCAT(Digest,TO_STRING(Hs[i],'{0:x8}')); END_FOR;
        Busy := FALSE; Done := TRUE; EXIT;
    END_IF;
END_FOR;
END_FUNCTION_BLOCK

(* ---- NG_Store.st ---- *)
FUNCTION_BLOCK NG_Store
VAR_INPUT
    Save : BOOL;
END_VAR
VAR_IN_OUT
    Candidate : NG_Durable;
END_VAR
VAR_OUTPUT
    Ready : BOOL;
    NeedsMigration : BOOL;
    Busy : BOOL;
    Done : BOOL;
    Error : BOOL;
    ErrorText : NG_Text;
    Active : NG_Durable;
END_VAR
VAR
    LegacyRecord : NG1_File;
    V2Record : NG2_File;
    V3Record : NG3_File;
    V4Record : NG4_File;
    V4 : BOOL;
    V3 : BOOL;
    V2 : BOOL;
    Legacy : BOOL;
    StateLength : UDINT;
    d : INT;
    p : INT;
    idx : INT;
    Stage : INT;
    Slot : INT := 1;
    ActiveSlot : INT;
    Prev : BOOL;
    Name : STRING;
    OpenFile : FILE_OPEN;
    ReadFile : FILE_READ;
    WriteFile : FILE_WRITE;
    CloseFile : FILE_CLOSE;
    Handle : UINT;
    Record : NG_File;
    Verify : NG_File;
    Bytes : NG_StorageBytes;
    CopyBytes : BUF_TO_BYTE;
    Hash : NG_StorageHash;
    Valid : BOOL;
    Saving : BOOL;
    OperationFailed : BOOL;
END_VAR
Done := FALSE;
IF Legacy THEN
    IF Slot = 1 THEN Name := '/opt/plcnext/NativeGateway-A.bin'; ELSE Name := '/opt/plcnext/NativeGateway-B.bin'; END_IF;
    StateLength := SIZEOF(LegacyRecord.State);
ELSIF V2 THEN
    IF Slot = 1 THEN Name := '/opt/plcnext/NativeGateway-v2-A.bin'; ELSE Name := '/opt/plcnext/NativeGateway-v2-B.bin'; END_IF;
    StateLength := SIZEOF(V2Record.State);
ELSIF V3 THEN
    IF Slot = 1 THEN Name := '/opt/plcnext/NativeGateway-v3-A.bin'; ELSE Name := '/opt/plcnext/NativeGateway-v3-B.bin'; END_IF;
    StateLength := SIZEOF(V3Record.State);
ELSIF V4 THEN
    IF Slot = 1 THEN Name := '/opt/plcnext/NativeGateway-v4-A.bin'; ELSE Name := '/opt/plcnext/NativeGateway-v4-B.bin'; END_IF;
    StateLength := SIZEOF(V4Record.State);
ELSE
    IF Slot = 1 THEN Name := '/opt/plcnext/NativeGateway-v5-A.bin'; ELSE Name := '/opt/plcnext/NativeGateway-v5-B.bin'; END_IF;
    StateLength := SIZEOF(Record.State);
END_IF;
OpenFile(Execute := (Stage = 10) OR (Stage = 60) OR (Stage = 90), Name := Name);
IF Legacy THEN
    ReadFile(Execute := Stage = 20, Handle := Handle, MaxLength := SIZEOF(LegacyRecord), Buffer := LegacyRecord);
ELSIF V2 THEN
    ReadFile(Execute := Stage = 20, Handle := Handle, MaxLength := SIZEOF(V2Record), Buffer := V2Record);
ELSIF V3 THEN
    ReadFile(Execute := Stage = 20, Handle := Handle, MaxLength := SIZEOF(V3Record), Buffer := V3Record);
ELSIF V4 THEN
    ReadFile(Execute := Stage = 20, Handle := Handle, MaxLength := SIZEOF(V4Record), Buffer := V4Record);
ELSE
    ReadFile(Execute := (Stage = 20) OR (Stage = 100), Handle := Handle, MaxLength := SIZEOF(Record), Buffer := Record);
END_IF;
WriteFile(Execute := Stage = 70, Handle := Handle, Length := SIZEOF(Record), Buffer := Record);
CloseFile(Execute := (Stage = 30) OR (Stage = 80) OR (Stage = 110) OR (Stage = 900), Handle := Handle);
IF Legacy THEN
    CopyBytes(REQ := Stage = 35, BUF_FORMAT := FALSE, BUF_OFFS := 0, BUF_CNT := StateLength, BUFFER := LegacyRecord.State, DST := Bytes);
ELSIF V2 THEN
    CopyBytes(REQ := Stage = 35, BUF_FORMAT := FALSE, BUF_OFFS := 0, BUF_CNT := StateLength, BUFFER := V2Record.State, DST := Bytes);
ELSIF V3 THEN
    CopyBytes(REQ := Stage = 35, BUF_FORMAT := FALSE, BUF_OFFS := 0, BUF_CNT := StateLength, BUFFER := V3Record.State, DST := Bytes);
ELSIF V4 THEN
    CopyBytes(REQ := Stage = 35, BUF_FORMAT := FALSE, BUF_OFFS := 0, BUF_CNT := StateLength, BUFFER := V4Record.State, DST := Bytes);
ELSE
    CopyBytes(REQ := (Stage = 35) OR (Stage = 50) OR (Stage = 115), BUF_FORMAT := FALSE, BUF_OFFS := 0, BUF_CNT := StateLength, BUFFER := Record.State, DST := Bytes);
END_IF;
Hash(Execute := (Stage = 40) OR (Stage = 55) OR (Stage = 120), Length := StateLength, Buffer := Bytes);
CASE Stage OF
0: Ready := FALSE; Busy := TRUE; Slot := 1; Stage := 10;
10:
    IF OpenFile.Error THEN Stage := 45;
    ELSIF OpenFile.Done THEN Handle := OpenFile.Handle; Stage := 20;
    END_IF;
20:
    IF ReadFile.Error OR ReadFile.Done THEN
        IF Legacy THEN Valid := ReadFile.Done AND (ReadFile.LengthRead = SIZEOF(LegacyRecord)) AND (LegacyRecord.Magic = DWORD#16#4E475731) AND (LegacyRecord.FormatVersion = 1);
        ELSIF V2 THEN Valid := ReadFile.Done AND (ReadFile.LengthRead = SIZEOF(V2Record)) AND (V2Record.Magic = DWORD#16#4E475732) AND (V2Record.FormatVersion = 2);
        ELSIF V3 THEN Valid := ReadFile.Done AND (ReadFile.LengthRead = SIZEOF(V3Record)) AND (V3Record.Magic = DWORD#16#4E475733) AND (V3Record.FormatVersion = 3);
        ELSIF V4 THEN Valid := ReadFile.Done AND (ReadFile.LengthRead = SIZEOF(V4Record)) AND (V4Record.Magic = DWORD#16#4E475734) AND (V4Record.FormatVersion = 4);
        ELSE Valid := ReadFile.Done AND (ReadFile.LengthRead = SIZEOF(Record)) AND (Record.Magic = DWORD#16#4E475735) AND (Record.FormatVersion = 5); END_IF;
        Stage := 30;
    END_IF;
30:
    IF CloseFile.Done OR CloseFile.Error THEN
        IF Valid AND NOT CloseFile.Error THEN Stage := 35; ELSE Stage := 45; END_IF;
    END_IF;
35: IF CopyBytes.DONE THEN Stage := 40; ELSIF CopyBytes.ERROR THEN Stage := 45; END_IF;
40:
    IF Hash.Done THEN
        IF Legacy THEN
            IF (Hash.Digest = LegacyRecord.Digest) AND (LegacyRecord.State.Generation > Active.Generation) THEN
                Active.Managed := FALSE; Active.BootCounter := 0;
                Active.Generation := LegacyRecord.State.Generation; Active.Bootstrap := LegacyRecord.State.Bootstrap;
                Active.ReplayIndex := LegacyRecord.State.ReplayIndex; Active.Requests := LegacyRecord.State.Requests;
                Active.Config.Version := LegacyRecord.State.Config.Version; Active.Config.MessageId := LegacyRecord.State.Config.MessageId;
                Active.Config.enabled := LegacyRecord.State.Config.enabled; Active.Config.batchIntervalMs := LegacyRecord.State.Config.batchIntervalMs;
                Active.Config.maxBatchPoints := LegacyRecord.State.Config.maxBatchPoints; Active.Config.DeviceCount := LegacyRecord.State.Config.DeviceCount;
                idx := 1;
                FOR d := 1 TO Active.Config.DeviceCount DO
                    Active.Config.Devices[d].deviceId := LegacyRecord.State.Config.Devices[d].deviceId;
                    Active.Config.Devices[d].name := LegacyRecord.State.Config.Devices[d].name;
                    Active.Config.Devices[d].enabled := LegacyRecord.State.Config.Devices[d].enabled;
                    Active.Config.Devices[d].host := LegacyRecord.State.Config.Devices[d].host;
                    Active.Config.Devices[d].port := LegacyRecord.State.Config.Devices[d].port;
                    Active.Config.Devices[d].unitId := LegacyRecord.State.Config.Devices[d].unitId;
                    Active.Config.Devices[d].connectTimeoutMs := LegacyRecord.State.Config.Devices[d].connectTimeoutMs;
                    Active.Config.Devices[d].requestTimeoutMs := LegacyRecord.State.Config.Devices[d].requestTimeoutMs;
                    Active.Config.Devices[d].retryCount := LegacyRecord.State.Config.Devices[d].retryCount;
                    Active.Config.Devices[d].maxReadRegisters := UINT#0;
                    Active.Config.Devices[d].hasMaxRegisterGap := FALSE;
                    Active.Config.Devices[d].maxRegisterGap := UINT#0;
                    Active.Config.Devices[d].PointCount := LegacyRecord.State.Config.Devices[d].PointCount;
                    Active.Config.Devices[d].PointStart := idx;
                    FOR p := 1 TO Active.Config.Devices[d].PointCount DO Active.Config.Points[idx] := LegacyRecord.State.Config.Devices[d].Points[p]; idx := idx+1; END_FOR;
                END_FOR;
                Active.Config.PointCount := idx-1; NeedsMigration := TRUE;
            END_IF;
        ELSIF V2 THEN
            IF (Hash.Digest = V2Record.Digest) AND (V2Record.State.Generation > Active.Generation) THEN
                Active.Generation := V2Record.State.Generation; Active.Bootstrap := V2Record.State.Bootstrap;
                Active.Config.Version := V2Record.State.Config.Version; Active.Config.MessageId := V2Record.State.Config.MessageId;
                Active.Config.enabled := V2Record.State.Config.enabled; Active.Config.batchIntervalMs := V2Record.State.Config.batchIntervalMs;
                Active.Config.maxBatchPoints := V2Record.State.Config.maxBatchPoints; Active.Config.DeviceCount := V2Record.State.Config.DeviceCount;
                Active.Config.PointCount := V2Record.State.Config.PointCount; Active.Config.Points := V2Record.State.Config.Points;
                FOR d := 1 TO Active.Config.DeviceCount DO
                    Active.Config.Devices[d].deviceId := V2Record.State.Config.Devices[d].deviceId; Active.Config.Devices[d].name := V2Record.State.Config.Devices[d].name;
                    Active.Config.Devices[d].enabled := V2Record.State.Config.Devices[d].enabled; Active.Config.Devices[d].host := V2Record.State.Config.Devices[d].host;
                    Active.Config.Devices[d].port := V2Record.State.Config.Devices[d].port; Active.Config.Devices[d].unitId := V2Record.State.Config.Devices[d].unitId;
                    Active.Config.Devices[d].connectTimeoutMs := V2Record.State.Config.Devices[d].connectTimeoutMs; Active.Config.Devices[d].requestTimeoutMs := V2Record.State.Config.Devices[d].requestTimeoutMs;
                    Active.Config.Devices[d].retryCount := V2Record.State.Config.Devices[d].retryCount;
                    Active.Config.Devices[d].maxReadRegisters := UINT#0; Active.Config.Devices[d].hasMaxRegisterGap := FALSE; Active.Config.Devices[d].maxRegisterGap := UINT#0;
                    Active.Config.Devices[d].PointCount := V2Record.State.Config.Devices[d].PointCount; Active.Config.Devices[d].PointStart := V2Record.State.Config.Devices[d].PointStart;
                END_FOR;
                Active.Requests := V2Record.State.Requests; Active.ReplayIndex := V2Record.State.ReplayIndex;
                Active.Managed := FALSE; Active.BootCounter := 0; NeedsMigration := TRUE;
            END_IF;
        ELSIF V3 THEN
            IF (Hash.Digest = V3Record.Digest) AND (V3Record.State.Generation > Active.Generation) THEN
                Active.Generation := V3Record.State.Generation; Active.Managed := V3Record.State.Managed;
                Active.BootCounter := V3Record.State.BootCounter; Active.Bootstrap := V3Record.State.Bootstrap;
                Active.Config.Version := V3Record.State.Config.Version; Active.Config.MessageId := V3Record.State.Config.MessageId;
                Active.Config.enabled := V3Record.State.Config.enabled; Active.Config.batchIntervalMs := V3Record.State.Config.batchIntervalMs;
                Active.Config.maxBatchPoints := V3Record.State.Config.maxBatchPoints; Active.Config.DeviceCount := V3Record.State.Config.DeviceCount;
                Active.Config.PointCount := V3Record.State.Config.PointCount; Active.Config.Points := V3Record.State.Config.Points;
                FOR d := 1 TO Active.Config.DeviceCount DO
                    Active.Config.Devices[d].deviceId := V3Record.State.Config.Devices[d].deviceId; Active.Config.Devices[d].name := V3Record.State.Config.Devices[d].name;
                    Active.Config.Devices[d].enabled := V3Record.State.Config.Devices[d].enabled; Active.Config.Devices[d].host := V3Record.State.Config.Devices[d].host;
                    Active.Config.Devices[d].port := V3Record.State.Config.Devices[d].port; Active.Config.Devices[d].unitId := V3Record.State.Config.Devices[d].unitId;
                    Active.Config.Devices[d].connectTimeoutMs := V3Record.State.Config.Devices[d].connectTimeoutMs; Active.Config.Devices[d].requestTimeoutMs := V3Record.State.Config.Devices[d].requestTimeoutMs;
                    Active.Config.Devices[d].retryCount := V3Record.State.Config.Devices[d].retryCount;
                    Active.Config.Devices[d].maxReadRegisters := UINT#0; Active.Config.Devices[d].hasMaxRegisterGap := FALSE; Active.Config.Devices[d].maxRegisterGap := UINT#0;
                    Active.Config.Devices[d].PointCount := V3Record.State.Config.Devices[d].PointCount; Active.Config.Devices[d].PointStart := V3Record.State.Config.Devices[d].PointStart;
                END_FOR;
                Active.Requests := V3Record.State.Requests; Active.ReplayIndex := V3Record.State.ReplayIndex;
                Active.HasHubBaseline := Active.Managed AND (Active.Config.Version > 0);
                IF Active.HasHubBaseline THEN Active.HubConfig := Active.Config; END_IF;
                Active.LocalChanges := FALSE; Active.LocalRevision := 0; NeedsMigration := TRUE;
            END_IF;
        ELSIF V4 THEN
            IF (Hash.Digest = V4Record.Digest) AND (V4Record.State.Generation > Active.Generation) THEN
                Active.Generation := V4Record.State.Generation; Active.Managed := V4Record.State.Managed;
                Active.BootCounter := V4Record.State.BootCounter; Active.Bootstrap := V4Record.State.Bootstrap;
                Active.HasHubBaseline := V4Record.State.HasHubBaseline; Active.LocalChanges := V4Record.State.LocalChanges; Active.LocalRevision := V4Record.State.LocalRevision;
                Active.Config.Version := V4Record.State.Config.Version; Active.Config.MessageId := V4Record.State.Config.MessageId;
                Active.Config.enabled := V4Record.State.Config.enabled; Active.Config.batchIntervalMs := V4Record.State.Config.batchIntervalMs;
                Active.Config.maxBatchPoints := V4Record.State.Config.maxBatchPoints; Active.Config.DeviceCount := V4Record.State.Config.DeviceCount;
                Active.Config.PointCount := V4Record.State.Config.PointCount; Active.Config.Points := V4Record.State.Config.Points;
                FOR d := 1 TO Active.Config.DeviceCount DO
                    Active.Config.Devices[d].deviceId := V4Record.State.Config.Devices[d].deviceId; Active.Config.Devices[d].name := V4Record.State.Config.Devices[d].name;
                    Active.Config.Devices[d].enabled := V4Record.State.Config.Devices[d].enabled; Active.Config.Devices[d].host := V4Record.State.Config.Devices[d].host;
                    Active.Config.Devices[d].port := V4Record.State.Config.Devices[d].port; Active.Config.Devices[d].unitId := V4Record.State.Config.Devices[d].unitId;
                    Active.Config.Devices[d].connectTimeoutMs := V4Record.State.Config.Devices[d].connectTimeoutMs; Active.Config.Devices[d].requestTimeoutMs := V4Record.State.Config.Devices[d].requestTimeoutMs;
                    Active.Config.Devices[d].retryCount := V4Record.State.Config.Devices[d].retryCount;
                    Active.Config.Devices[d].maxReadRegisters := UINT#0; Active.Config.Devices[d].hasMaxRegisterGap := FALSE; Active.Config.Devices[d].maxRegisterGap := UINT#0;
                    Active.Config.Devices[d].PointCount := V4Record.State.Config.Devices[d].PointCount; Active.Config.Devices[d].PointStart := V4Record.State.Config.Devices[d].PointStart;
                END_FOR;
                Active.HubConfig.Version := V4Record.State.HubConfig.Version; Active.HubConfig.MessageId := V4Record.State.HubConfig.MessageId;
                Active.HubConfig.enabled := V4Record.State.HubConfig.enabled; Active.HubConfig.batchIntervalMs := V4Record.State.HubConfig.batchIntervalMs;
                Active.HubConfig.maxBatchPoints := V4Record.State.HubConfig.maxBatchPoints; Active.HubConfig.DeviceCount := V4Record.State.HubConfig.DeviceCount;
                Active.HubConfig.PointCount := V4Record.State.HubConfig.PointCount; Active.HubConfig.Points := V4Record.State.HubConfig.Points;
                FOR d := 1 TO Active.HubConfig.DeviceCount DO
                    Active.HubConfig.Devices[d].deviceId := V4Record.State.HubConfig.Devices[d].deviceId; Active.HubConfig.Devices[d].name := V4Record.State.HubConfig.Devices[d].name;
                    Active.HubConfig.Devices[d].enabled := V4Record.State.HubConfig.Devices[d].enabled; Active.HubConfig.Devices[d].host := V4Record.State.HubConfig.Devices[d].host;
                    Active.HubConfig.Devices[d].port := V4Record.State.HubConfig.Devices[d].port; Active.HubConfig.Devices[d].unitId := V4Record.State.HubConfig.Devices[d].unitId;
                    Active.HubConfig.Devices[d].connectTimeoutMs := V4Record.State.HubConfig.Devices[d].connectTimeoutMs; Active.HubConfig.Devices[d].requestTimeoutMs := V4Record.State.HubConfig.Devices[d].requestTimeoutMs;
                    Active.HubConfig.Devices[d].retryCount := V4Record.State.HubConfig.Devices[d].retryCount;
                    Active.HubConfig.Devices[d].maxReadRegisters := UINT#0; Active.HubConfig.Devices[d].hasMaxRegisterGap := FALSE; Active.HubConfig.Devices[d].maxRegisterGap := UINT#0;
                    Active.HubConfig.Devices[d].PointCount := V4Record.State.HubConfig.Devices[d].PointCount; Active.HubConfig.Devices[d].PointStart := V4Record.State.HubConfig.Devices[d].PointStart;
                END_FOR;
                Active.Requests := V4Record.State.Requests; Active.ReplayIndex := V4Record.State.ReplayIndex;
                NeedsMigration := TRUE;
            END_IF;
        ELSIF (Hash.Digest = Record.Digest) AND (Record.State.Generation > Active.Generation) THEN Active := Record.State; ActiveSlot := Slot; END_IF;
        Stage := 45;
    END_IF;
45:
    IF Slot = 1 THEN Slot := 2; Stage := 10;
    ELSIF (Active.Generation = 0) AND NOT Legacy AND NOT V2 AND NOT V3 AND NOT V4 THEN V4 := TRUE; Slot := 1; Stage := 10;
    ELSIF (Active.Generation = 0) AND V4 THEN V4 := FALSE; V3 := TRUE; Slot := 1; Stage := 10;
    ELSIF (Active.Generation = 0) AND V3 THEN V3 := FALSE; V2 := TRUE; Slot := 1; Stage := 10;
    ELSIF (Active.Generation = 0) AND V2 THEN V2 := FALSE; Legacy := TRUE; Slot := 1; Stage := 10;
    ELSE Ready := TRUE; Busy := FALSE; Stage := 200; END_IF;
50: IF CopyBytes.DONE THEN Stage := 55; ELSIF CopyBytes.ERROR THEN Error := TRUE; ErrorText := 'STORAGE_ERROR'; Busy := FALSE; Stage := 200; END_IF;
55:
    IF Hash.Done THEN Record.Digest := Hash.Digest; Stage := 60; END_IF;
60:
    IF OpenFile.Error THEN Error := TRUE; ErrorText := 'STORAGE_ERROR'; Busy := FALSE; Stage := 200;
    ELSIF OpenFile.Done THEN Handle := OpenFile.Handle; Stage := 70; END_IF;
70:
    IF WriteFile.Error OR WriteFile.Done THEN
        OperationFailed := WriteFile.Error OR (WriteFile.LengthWritten <> SIZEOF(Record)); Stage := 80;
    END_IF;
80:
    IF CloseFile.Done OR CloseFile.Error THEN
        IF OperationFailed OR CloseFile.Error THEN Error := TRUE; ErrorText := 'STORAGE_ERROR'; Busy := FALSE; Stage := 200;
        ELSE Verify := Record; Stage := 85; END_IF;
    END_IF;
85: Stage := 90;
90:
    IF OpenFile.Error THEN Error := TRUE; ErrorText := 'STORAGE_ERROR'; Busy := FALSE; Stage := 200;
    ELSIF OpenFile.Done THEN Handle := OpenFile.Handle; Stage := 100; END_IF;
100:
    IF ReadFile.Error OR ReadFile.Done THEN
        Valid := ReadFile.Done AND (ReadFile.LengthRead = SIZEOF(Record)) AND (Record.Magic = Verify.Magic) AND (Record.FormatVersion = 5) AND (Record.State.Generation = Verify.State.Generation);
        Stage := 110;
    END_IF;
110:
    IF CloseFile.Done OR CloseFile.Error THEN
        IF Valid AND NOT CloseFile.Error THEN Stage := 115;
        ELSE Error := TRUE; ErrorText := 'STORAGE_ERROR'; Busy := FALSE; Stage := 200; END_IF;
    END_IF;
115: IF CopyBytes.DONE THEN Stage := 120; ELSIF CopyBytes.ERROR THEN Error := TRUE; ErrorText := 'STORAGE_ERROR'; Busy := FALSE; Stage := 200; END_IF;
120:
    IF Hash.Done THEN
        IF (Hash.Digest = Verify.Digest) AND (Record.Digest = Verify.Digest) THEN
            Active := Record.State; ActiveSlot := Slot; Done := TRUE; NeedsMigration := FALSE;
        ELSE Error := TRUE; ErrorText := 'STORAGE_ERROR'; END_IF;
        Busy := FALSE; Stage := 200;
    END_IF;
200:
    IF Save AND NOT Prev THEN
        Error := FALSE; ErrorText := ''; Busy := TRUE;
        Legacy := FALSE; V2 := FALSE; V3 := FALSE; V4 := FALSE;
        Record.Magic := DWORD#16#4E475735; Record.FormatVersion := 5;
        Record.State := Candidate; Record.State.Generation := Active.Generation+1;
        IF ActiveSlot = 1 THEN Slot := 2; ELSE Slot := 1; END_IF;
        Stage := 50;
    END_IF;
END_CASE;
Prev := Save;
END_FUNCTION_BLOCK
